(* IEC 61131-3 sources: RootPLC/blocks/templates/filling-station, 2 files *)

(* ---- filling_station.st ---- *)
(* L4 template: filling station (blocks/templates/filling-station/README.md).
   Containers are filled with a timed dose from a buffer tank; the tank's
   level is held by an inlet valve. Built only from RootBlocks blocks
   (--library RootBlocks). No I/O inside: io_map.st binds it to the board. *)
FUNCTION_BLOCK FB_FillingStation
VAR_INPUT
    (* operator *)
    ReqOff           : BOOL;
    ReqManual        : BOOL;
    ReqAuto          : BOOL;
    StartBtn         : BOOL;
    StopBtn          : BOOL;
    ResetBtn         : BOOL;            (* also acknowledges alarms *)
    ManInlet         : BOOL;            (* manual commands *)
    ManPump          : BOOL;
    EStopOk          : BOOL := TRUE;    (* status from the safety relay *)
    (* plant *)
    LevelRaw         : REAL;            (* level transmitter, 0 .. 27648 *)
    HighLevelSw      : BOOL;            (* TRUE: tank level high *)
    LowLevelSw       : BOOL;            (* TRUE: enough liquid for the pump *)
    InletOpenFb      : BOOL;
    InletClosedFb    : BOOL;
    PumpRunningFb    : BOOL;
    PumpOverload     : BOOL;
    ContainerPresent : BOOL;
    (* parameters *)
    LevelSP          : REAL := 60.0;    (* % *)
    LevelBand        : REAL := 20.0;    (* % *)
    DoseTime         : TIME := T#3s;
    BatchSize        : UDINT := 10;
END_VAR
VAR_OUTPUT
    InletValve  : BOOL;
    Pump        : BOOL;
    LampRunning : BOOL;
    LampFault   : BOOL;
    LampAlarm   : BOOL;
    Level       : REAL;                 (* % *)
    Filled      : UDINT;                (* containers in this batch *)
    State       : RB_MACHINE_STATE;
    Mode        : RB_MODE;
END_VAR
VAR
    modes     : RB_ModeManager;
    machine   : RB_MachineState;
    levelIn   : RB_Scale;
    levelPv   : RB_FilterPT1;
    levelCtl  : RB_OnOff;
    inlet     : RB_ValveOnOff;
    pumpDev   : RB_Pump;
    container : RB_Debounce;
    chain     : RB_StepChain;
    highAlarm : RB_Alarm;
    count     : RB_Counter;
    fault     : BOOL;
    running   : BOOL;
    aborted   : BOOL;
    proceed   : BOOL;
END_VAR

(* devices and measurements report faults; any fault aborts the machine *)
fault := inlet.Error OR pumpDev.Error OR levelIn.Error;
modes(ReqOff := ReqOff, ReqManual := ReqManual, ReqAuto := ReqAuto,
      EStopOk := EStopOk, Fault := fault);
Mode := modes.Mode;

(* the reset button clears an abort, otherwise it resets the machine *)
aborted := machine.State = RB_MACHINE_STATE#Aborted;
machine(Reset := ResetBtn AND NOT aborted, Clear := ResetBtn AND aborted,
        Start := StartBtn AND Mode = RB_MODE#Auto,
        Stop := StopBtn OR Mode <> RB_MODE#Auto OR count.Done,
        Abort := NOT EStopOk OR fault,
        ResetDone := NOT fault, StartDone := TRUE,
        StopDone := chain.StepNo <= 1);
State := machine.State;
running := State = RB_MACHINE_STATE#Execute OR State = RB_MACHINE_STATE#Stopping;

(* level: scale, smooth, hold between SP - band/2 and SP + band/2; the
   inlet follows it in Auto, and a high level closes it in every mode *)
levelIn(Raw := LevelRaw, RawMin := 0.0, RawMax := 27648.0, EngMin := 0.0, EngMax := 100.0,
        Margin := 500.0, Reset := ResetBtn);
levelPv(In := levelIn.Value, T := T#500ms);
Level := levelPv.Out;
levelCtl(Enable := TRUE, SP := LevelSP, PV := Level, Hysteresis := LevelBand);
highAlarm(In := HighLevelSw, OnDelay := T#1s, Ack := ResetBtn);
inlet(Mode := Mode, AutoOpen := levelCtl.Out, ManOpen := ManInlet, Interlock := HighLevelSw,
      FbOpen := InletOpenFb, FbClosed := InletClosedFb, Reset := ResetBtn);

(* one container, a cyclic chain: 1 wait for it, 2 dose, 3 wait until it
   is taken away, then 1 again *)
container(In := ContainerPresent, OnDelay := T#200ms, OffDelay := T#200ms);
CASE chain.StepNo OF
1: proceed := container.Out AND State = RB_MACHINE_STATE#Execute;
2: proceed := chain.StepTime >= DoseTime;
3: proceed := NOT container.Out;
END_CASE;
chain(Start := running, Proceed := proceed, NextStep := chain.StepNo MOD 3 + 1,
      Abort := NOT running);
pumpDev(Mode := Mode, AutoRun := chain.StepNo = 2, ManRun := ManPump,
        FbRunning := PumpRunningFb, Overload := PumpOverload, DryRun := NOT LowLevelSw,
        DryRunTime := T#1s, Reset := ResetBtn);
count(In := chain.StepNo = 3, Preset := BatchSize,
      Reset := State = RB_MACHINE_STATE#Starting);
Filled := count.Count;

InletValve := inlet.Open;
Pump := pumpDev.Run;
LampRunning := machine.Producing;
LampFault := fault OR State = RB_MACHINE_STATE#Aborted;
LampAlarm := highAlarm.Active OR highAlarm.Unacked;
END_FUNCTION_BLOCK

(* ---- io_map.st ---- *)
(* The filling station on a controller: located I/O bound to the template
   (spec/14-runtime.md). Adapt the addresses to the board's I/O modules.
   Run: rootplc runtime blocks/templates/filling-station --library RootBlocks
        --program PLC_PRG --modbus 5502 *)
PROGRAM PLC_PRG
VAR
    (* digital inputs *)
    btnAuto       AT %IX0.0 : BOOL;
    btnManual     AT %IX0.1 : BOOL;
    btnOff        AT %IX0.2 : BOOL;
    btnStart      AT %IX0.3 : BOOL;
    btnStop       AT %IX0.4 : BOOL;
    btnReset      AT %IX0.5 : BOOL;
    estopOk       AT %IX0.6 : BOOL;
    highLevel     AT %IX0.7 : BOOL;
    lowLevel      AT %IX1.0 : BOOL;
    inletOpen     AT %IX1.1 : BOOL;
    inletClosed   AT %IX1.2 : BOOL;
    pumpRunning   AT %IX1.3 : BOOL;
    pumpOverload  AT %IX1.4 : BOOL;
    containerIn   AT %IX1.5 : BOOL;
    (* analog input *)
    levelRaw      AT %IW2 : INT;
    (* manual commands from the HMI (Modbus holding register 0) *)
    hmiManual     AT %MW0 : WORD;
    (* outputs *)
    inletValve    AT %QX0.0 : BOOL;
    pump          AT %QX0.1 : BOOL;
    lampRunning   AT %QX0.2 : BOOL;
    lampFault     AT %QX0.3 : BOOL;
    lampAlarm     AT %QX0.4 : BOOL;
    levelPercent  AT %QW2 : INT;    (* level in 0.1 % for the HMI *)
    filledCount   AT %QW4 : UINT;
    station       : FB_FillingStation;
END_VAR
station(ReqAuto := btnAuto, ReqManual := btnManual, ReqOff := btnOff,
        StartBtn := btnStart, StopBtn := btnStop, ResetBtn := btnReset,
        ManInlet := (hmiManual AND WORD#1) <> WORD#0,
        ManPump := (hmiManual AND WORD#2) <> WORD#0,
        EStopOk := estopOk, LevelRaw := INT_TO_REAL(levelRaw),
        HighLevelSw := highLevel, LowLevelSw := lowLevel,
        InletOpenFb := inletOpen, InletClosedFb := inletClosed,
        PumpRunningFb := pumpRunning, PumpOverload := pumpOverload,
        ContainerPresent := containerIn);
inletValve := station.InletValve;
pump := station.Pump;
lampRunning := station.LampRunning;
lampFault := station.LampFault;
lampAlarm := station.LampAlarm;
levelPercent := REAL_TO_INT(station.Level * 10.0);
filledCount := UDINT_TO_UINT(station.Filled);
END_PROGRAM
